ORGANIZATION_BLOCK
BEGIN
END_ORGANIZATION_BLOCK
